(* IEC 61131-3 sources: axsharp/src/ix.templates/working/templates/ixtwin/ax/src, 2 files *)

(* ---- configuration.st ---- *)
CONFIGURATION MyConfiguration
    TASK Main(Interval := T#10ms, Priority := 1);
    PROGRAM P1 WITH Main: MainProgram;

    VAR_GLOBAL

    END_VAR
END_CONFIGURATION

(* ---- program.st ---- *)
PROGRAM MainProgram
    VAR_EXTERNAL

    END_VAR

    VAR

    END_VAR

    VAR_TEMP

    END_VAR

    // code here
    ;
END_PROGRAM
